// TIA Portal V21 export
// export: Created 2026-11-11T00:49:01.4904174Z, ExportSetting WithDefaults, DisplayName Totally Integrated Automation Portal, DisplayVersion V21 Update 3, DisplayName STEP 7 Professional, DisplayVersion V21 Update 3, DisplayName STEP 7 Safety, DisplayVersion V21, DisplayName Tech WebApplication, DisplayVersion V21, DisplayName WinCC Basic/Comfort/Advanced, DisplayVersion V21 Update 3, DisplayName WinCC Unified, DisplayVersion V21 Update 3
FUNCTION_BLOCK "FX_Lad_ex070"   // FB257, LAD
{ S7_Optimized_Access := 'TRUE' }
VERSION : 0.1
// stored: AutoNumber true, IsIECCheckEnabled false, IsRetainMemResEnabled false, MemoryReserve 100, SetENOAutomatically false, UDAEnableTagReadback false
   VAR_INPUT
      "a" : Bool;
      "b" : Bool;
      c : Bool;
      ia : Int;
      ib : Int;
      ic : Int;
      da : DInt;
      db : DInt;
      ra : Real;
      rb : Real;
      wa : Word;
      wb : Word;
      dwa : DWord;
      ba : Byte;
      ta : Time;
      tb : Time;
      s1 : String;
      s2 : String;
   END_VAR
   VAR_OUTPUT
      q : Bool;
      q2 : Bool;
      io : Int;
      io2 : Int;
      dout : DInt;
      rout : Real;
      wout : Word;
      dwout : DWord;
      bout : Byte;
      tout : Time;
      sout : String;
   END_VAR
   VAR_IN_OUT
      p_enable : Bool;
      p_id : HW_SUBMODULE;
      p_slot_no_x : Int;
      p_func_x : Int;
      p_busy : Bool;
      p_done : Bool;
      p_error : Bool;
      p_status : DWord;
      x_int : Int;
      arr : Array[0..9] of Int;
      barr : Array[0..7] of Bool;
      iinout : Int;
   END_VAR
   VAR
      inst : PE_DS3_Write_ET200S;
      ton1 { S7_SetPoint := 'True'} : TON_TIME;
      tof1 { S7_SetPoint := 'True'} : TOF_TIME;
      tp1 { S7_SetPoint := 'True'} : TP_TIME;
      tonr1 { S7_SetPoint := 'True'} : TONR_TIME;
      ctu1 { S7_SetPoint := 'True'} : CTU_INT;
      ctd1 { S7_SetPoint := 'True'} : CTD_INT;
      ctud1 { S7_SetPoint := 'True'} : CTUD_INT;
      rtrig1 { S7_SetPoint := 'True'} : R_TRIG;
      ftrig1 { S7_SetPoint := 'True'} : F_TRIG;
      edge1 : Bool;
      edge2 : Bool;
      stat1 : Bool;
      stat2 : Bool;
      stati : Int;
   END_VAR
   VAR_TEMP
      t1 : Bool;
      t2 : Bool;
      ti : Int;
      td : DInt;
      tr : Real;
      tw : Word;
      tt : Time;
      var1 : Variant;
   END_VAR
BEGIN

REGION Network 1: ---| |--- - Normally open contact
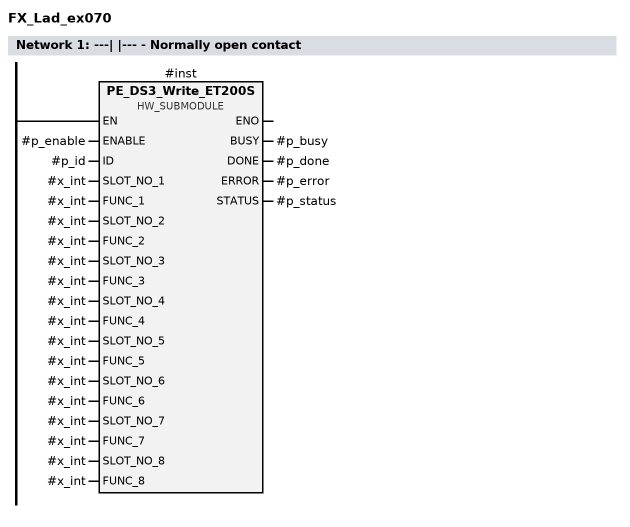
   RUNG wire#powerrail
      { S7_Templates := "id_type := HW_SUBMODULE" } #inst.PE_DS3_Write_ET200S(enable := #p_enable, ID := #p_id, busy => #p_busy, done => #p_done, error => #p_error, status => #p_status, Slot_No_1 := #x_int, Func_1 := #x_int, Slot_No_2 := #x_int, Func_2 := #x_int, Slot_No_3 := #x_int, Func_3 := #x_int, Slot_No_4 := #x_int, Func_4 := #x_int, Slot_No_5 := #x_int, Func_5 := #x_int, Slot_No_6 := #x_int, Func_6 := #x_int, Slot_No_7 := #x_int, Func_7 := #x_int, Slot_No_8 := #x_int, Func_8 := #x_int)
   END_RUNG
   // the same network as SCL:
   #inst(enable := #p_enable,   // PE_DS3_Write_ET200S
         ID := #p_id,
         Slot_No_1 := #x_int,
         Func_1 := #x_int,
         Slot_No_2 := #x_int,
         Func_2 := #x_int,
         Slot_No_3 := #x_int,
         Func_3 := #x_int,
         Slot_No_4 := #x_int,
         Func_4 := #x_int,
         Slot_No_5 := #x_int,
         Func_5 := #x_int,
         Slot_No_6 := #x_int,
         Func_6 := #x_int,
         Slot_No_7 := #x_int,
         Func_7 := #x_int,
         Slot_No_8 := #x_int,
         Func_8 := #x_int,
         busy => #p_busy,
         done => #p_done,
         error => #p_error,
         status => #p_status);
END_REGION
END_FUNCTION_BLOCK
